Fanuc KAREL source: kt00206.KL

-- PROVISIONAL review KL for V940-1; original PC SHA256 2ab6fbe3c9690139116cf6795750294425be311db75e5900560bb1328dc3a3ce
-- Incomplete behavior may be omitted. Consult companion uncertainty JSON. Do not deploy.
PROGRAM KT00206
%NOLOCKGROUP
VAR
  I1 : INTEGER
  OUT : INTEGER
-- UNRESOLVED_DECL Y2 type=002018
BEGIN
  -- V9_ZERO_TABLE_METADATA_HINT layout=0001; no indexed target words; source/name/runtime held
  -- UNRESOLVED_PC offsets 5-16; opcodes 2E,23
  -- UNRESOLVED_PC offsets 21-35; opcodes 2E,22,9D,33,B2
  -- UNRESOLVED_PC offsets 40-62; opcodes 21,22,9D,33,B1,46,23
  -- UNRESOLVED_PC offsets 67-71; opcodes 7F
END KT00206
